(* IEC 61131-3 sources: volt/packages/volt-lsp-iec/test-corpus/awa-palletizer/Device/Plc Logic/Application/Library Manager/L_SEMP_ErrorManagement, 51 files *)

(* ---- EVTPARAM_CMPLENZEERRORMANAGEMENTACCESSACTSTATEDETERMINEEVENTCHANGED.dut ---- *)
TYPE EVTPARAM_CMPLENZEERRORMANAGEMENTACCESSACTSTATEDETERMINEEVENTCHANGED :
STRUCT
	SEVERITY : USINT;
	EVENTID : WORD;
	TEXTREFID : WORD;
	ACTSTATEDETERMINEEVENT : DWORD;
END_STRUCT
END_TYPE

(* ---- EVTPARAM_CMPLENZEERRORMANAGEMENTACCESSACTSTATEDETERMINEEVENTCHANGED_V2.dut ---- *)
TYPE EVTPARAM_CMPLENZEERRORMANAGEMENTACCESSACTSTATEDETERMINEEVENTCHANGED_V2 :
STRUCT
	SEVERITY : USINT;
	EVENTID : WORD;
	TEXTREFID : WORD;
	ACTSTATEDETERMINEEVENT : DWORD;
	USERGROUP : WORD;
	USERPRIORITY : WORD;
	EVENTCONTROL : WORD;
END_STRUCT
END_TYPE

(* ---- EVTPARAM_CMPLENZEERRORMANAGEMENTACCESSCOMMANDEVENTREACTION.dut ---- *)
TYPE EVTPARAM_CMPLENZEERRORMANAGEMENTACCESSCOMMANDEVENTREACTION :
STRUCT
	SEVERITY : USINT;
	EVENTID : WORD;
	TEXTREFID : WORD;
END_STRUCT
END_TYPE

(* ---- EVTPARAM_CMPLENZEERRORMANAGEMENTACCESSRESETCOMPONENTOCCURRED.dut ---- *)
TYPE EVTPARAM_CMPLENZEERRORMANAGEMENTACCESSRESETCOMPONENTOCCURRED :
STRUCT
	INSTANCEID : UDINT;
	LAYER : USINT;
	SEVERITY : USINT;
	STATE : USINT;
	EVENTID : WORD;
	TEXTREFID : WORD;
END_STRUCT
END_TYPE

(* ---- EVTPARAM_CMPLENZEERRORMANAGEMENTACCESSRESETOCCURRED.dut ---- *)
TYPE EVTPARAM_CMPLENZEERRORMANAGEMENTACCESSRESETOCCURRED :
STRUCT
	ACTHIGHESTPRIOREVENT : POINTER TO L_SEMP_ActEvent;
	PCOMPLIST : POINTER TO L_SEMP_ComponentListResetOccured;
END_STRUCT
END_TYPE

(* ---- L_SEMP_ACTEVENT.dut ---- *)
TYPE L_SEMP_ACTEVENT :
STRUCT
	LAYER : USINT;
	SEVERITY : USINT;
	STATE : USINT;
	EVENTID : WORD;
	TEXTREFID : WORD;
	INSTANCEID : DWORD;
	ACTSTATEDETERMINEEVENT : DWORD;
	TIMESTAMP : L_SEMP_LogTimeStamp;
END_STRUCT
END_TYPE

(* ---- L_SEMP_BEHAVIOUR.dut ---- *)
TYPE L_SEMP_BEHAVIOUR :
(
	PROCESSERRORREACTION := 0,
	ONLYLOGGING := 1
);
END_TYPE

(* ---- L_SEMP_COMPONENTLISTRESETOCCURED.dut ---- *)
TYPE L_SEMP_COMPONENTLISTRESETOCCURED :
STRUCT
	PREVCMP : POINTER TO L_SEMP_ComponentListResetOccured;
	PCOMPONENT : POINTER TO DWORD;
	NEXTCMP : POINTER TO L_SEMP_ComponentListResetOccured;
END_STRUCT
END_TYPE

(* ---- L_SEMP_EVENTCONTROL.dut ---- *)
TYPE L_SEMP_EVENTCONTROL :
(
	NOACKNOLAGENEEDED := 0,
	ACKNOLAGENEEDED := 1,
	EVENTCONTROLNOTUSED := 255
);
END_TYPE

(* ---- L_SEMP_EVENTPARAMETERS.dut ---- *)
TYPE L_SEMP_EVENTPARAMETERS :
STRUCT
	EVENTPARAMETERS : ARRAY [1..10] OF L_SEMP_ParameterItem;
END_STRUCT
END_TYPE

(* ---- L_SEMP_EVENTPARAMETERSSHORT.dut ---- *)
TYPE L_SEMP_EVENTPARAMETERSSHORT :
STRUCT
	EVENTPARAMETERS : ARRAY [1..10] OF L_SEMP_ParameterItemShort;
END_STRUCT
END_TYPE

(* ---- L_SEMP_GROUP.dut ---- *)
TYPE L_SEMP_GROUP :
(
	USERGROUP1 := 1,
	USERGROUP2 := 2,
	USERGROUP3 := 3,
	USERGROUP4 := 4,
	USERGROUP5 := 5,
	MANUFACTURERGROUP1 := 11,
	MANUFACTURERGROUP2 := 12
);
END_TYPE

(* ---- L_SEMP_LAYER.dut ---- *)
TYPE L_SEMP_LAYER :
(
	KINEMATICS := 6,
	MOTION := 7,
	APPLICATION := 8,
	IEC_APPLICATION := 40,
	TA_LAYER := 50
);
END_TYPE

(* ---- L_SEMP_LAYER_INTERN.dut ---- *)
TYPE L_SEMP_LAYER_INTERN :
(
	LEM_LA_I900_BASE_FW := 0,
	LEM_LA_SAFETY := 1,
	LEM_LA_FEEDBACK := 2,
	LEM_LA_ETC_SLAVE := 3,
	LEM_LA_BASE_SETTINGS := 4,
	LEM_LA_COMMUNICATION := 5,
	LEM_LA_KINEMATICS := 6,
	LEM_LA_MOTION := 7,
	LEM_LA_TECH_APPLICATION := 8,
	LEM_LA_FIELDBUS := 10,
	LEM_LA_LEM := 20,
	LEM_LA_IEC_RUNTIME := 30,
	LEM_LA_ETC_MASTER := 31,
	LEM_LA_I900_IO_DRIVER := 32,
	LEM_LA_IEC_APPLICATION := 40,
	LEM_LA_TA_LAYER := 50
);
END_TYPE

(* ---- L_SEMP_LOGTIMESTAMP.dut ---- *)
TYPE L_SEMP_LOGTIMESTAMP :
STRUCT
	DWLOWDATETIME : DWORD;
	DWHIGHDATETIME : DWORD;
END_STRUCT
END_TYPE

(* ---- L_SEMP_PARAMETERITEM.dut ---- *)
TYPE L_SEMP_PARAMETERITEM :
STRUCT
	SIZE : BYTE;
	ETYPE : INT;
	VALUE : L_SEMP_ParaValue;
END_STRUCT
END_TYPE

(* ---- L_SEMP_PARAMETERITEMSHORT.dut ---- *)
TYPE L_SEMP_PARAMETERITEMSHORT :
STRUCT
	SIZE : BYTE;
	ETYPE : INT;
	VALUE : L_SEMP_ParaValueShort;
END_STRUCT
END_TYPE

(* ---- L_SEMP_PARAVALUE.dut ---- *)
TYPE L_SEMP_PARAVALUE :
UNION
	DWVALUE : DWORD;
	DNVALUE : DINT;
	FVALUE : REAL;
	STVALUE : STRING;
	DWTEXTLISTID : DWORD;
END_UNION
END_TYPE

(* ---- L_SEMP_PARAVALUESHORT.dut ---- *)
TYPE L_SEMP_PARAVALUESHORT :
UNION
	DWVALUE : DWORD;
	DNVALUE : DINT;
	RVALUE : REAL;
	LRVALUE : LREAL;
	DWTEXTLISTID : DWORD;
END_UNION
END_TYPE

(* ---- L_SEMP_PRIORITY.dut ---- *)
TYPE L_SEMP_PRIORITY :
(
	PRIORITY_1 := 1,
	PRIORITY_2 := 2,
	PRIORITY_3 := 3,
	PRIORITY_4 := 4,
	PRIORITY_5 := 5,
	PRIORITY_INFO_NOT_USED := 255
);
END_TYPE

(* ---- L_SEMP_SERVERITY.dut ---- *)
TYPE L_SEMP_SERVERITY :
(
	LEM_SEV_NO_RESPONSE := 0,
	LEM_SEV_FAULT_CIA402 := 1,
	LEM_SEV_WARNING := 2,
	LEM_SEV_INFORMATION := 11,
	LEM_SEV_WARNING_LOCK := 13,
	LEM_SEV_TROUBLE_LOG := 15,
	LEM_SEV_TROUBLE := 16,
	LEM_SEV_FAULT_LOG := 18,
	LEM_SEV_FAULT_FAST_STOP := 19,
	LEM_SEV_FAULT_QSP := 20,
	LEM_SEV_FAULT_CINH := 21,
	LEM_SEV_FAULT := 23
);
END_TYPE

(* ---- L_SEMP_SERVERITYLEVEL.dut ---- *)
TYPE L_SEMP_SERVERITYLEVEL :
(
	NO_RESPONSE := 0,
	FAULT_CIA402 := 1,
	WARNING := 2,
	INFORMATION := 11,
	WARNING_LOCK := 13,
	TROUBLE_LOG := 15,
	TROUBLE := 16,
	FAULT_FAST_STOP := 19,
	FAULT_QSP := 20,
	FAULT_QSP_CINH := 21,
	FAULT := 23
);
END_TYPE

(* ---- L_SEMP_EVENTIDS.gvl ---- *)
VAR_GLOBAL
	CMPID_CMPLENZEERRORMANAGEMENTACCESS : DWORD := 16#2014;
	EVT_CMPLENZEERRORMANAGEMENTACCESSACTSTATEDETERMINEEVENTCHANGED : DWORD := 16#10000011;
	EVTPARAMID_CMPLENZEERRORMANAGEMENTACCESSACTSTATEDETERMINEEVENTCHANGED : WORD := 16#1;
	EVTVERSION_CMPLENZEERRORMANAGEMENTACCESSACTSTATEDETERMINEEVENTCHANGED : WORD := 16#1;
	EVT_CMPLENZEERRORMANAGEMENTACCESSRESETOCCURRED : DWORD := 16#10000012;
	EVTPARAMID_CMPLENZEERRORMANAGEMENTACCESSRESETOCCURRED : WORD := 16#1;
	EVTVERSION_CMPLENZEERRORMANAGEMENTACCESSRESETOCCURRED : WORD := 16#1;
	EVT_CMPLENZEERRORMANAGEMENTACCESSCOMMANDEVENTREACTION : DWORD := 16#10000013;
	EVTPARAMID_CMPLENZEERRORMANAGEMENTACCESSCOMMANDEVENTREACTION : WORD := 16#1;
	EVTVERSION_CMPLENZEERRORMANAGEMENTACCESSCOMMANDEVENTREACTION : WORD := 16#1;
	EVT_CMPLENZEERRORMANAGEMENTACCESSREADACTERRORDATAAVAILABLE : DWORD := 16#10000014;
	EVTPARAMID_CMPLENZEERRORMANAGEMENTACCESSREADACTERRORDATAAVAILABLE : WORD := 16#1;
	EVTVERSION_CMPLENZEERRORMANAGEMENTACCESSREADACTERRORDATAAVAILABLE : WORD := 16#1;
END_VAR

(* ---- GETBOOLEANPROPERTY.pou ---- *)
FUNCTION GETBOOLEANPROPERTY : BOOL
VAR_INPUT
	STKEY : WSTRING;
END_VAR
END_FUNCTION

(* ---- GETCOMPANY.pou ---- *)
FUNCTION GETCOMPANY : WSTRING
END_FUNCTION

(* ---- GETNUMBERPROPERTY.pou ---- *)
FUNCTION GETNUMBERPROPERTY : DINT
VAR_INPUT
	STKEY : WSTRING;
END_VAR
END_FUNCTION

(* ---- GETTEXTPROPERTY.pou ---- *)
FUNCTION GETTEXTPROPERTY : WSTRING
VAR_INPUT
	STKEY : WSTRING;
END_VAR
END_FUNCTION

(* ---- GETTEXTPROPERTY2.pou ---- *)
FUNCTION GETTEXTPROPERTY2 : POINTER TO WSTRING
VAR_INPUT
	STKEY : WSTRING;
END_VAR
END_FUNCTION

(* ---- GETTITLE.pou ---- *)
FUNCTION GETTITLE : WSTRING
END_FUNCTION

(* ---- GETVERSION.pou ---- *)
FUNCTION GETVERSION : VERSION
END_FUNCTION

(* ---- GETVERSIONPROPERTY.pou ---- *)
FUNCTION GETVERSIONPROPERTY : VERSION
VAR_INPUT
	STKEY : WSTRING;
END_VAR
END_FUNCTION

(* ---- L_SEMP_CLEAREVENT.pou ---- *)
FUNCTION L_SEMP_CLEAREVENT : RTS_IEC_RESULT
VAR_INPUT
	HHANDLE : RTS_IEC_HANDLE := RTS_INVALID_HANDLE;
	UIEVENTID : UINT := 16#0;
END_VAR
END_FUNCTION

(* ---- L_SEMP_CLEAREVENT_V2.pou ---- *)
FUNCTION L_SEMP_CLEAREVENT_V2 : RTS_IEC_RESULT
VAR_INPUT
	HHANDLE : RTS_IEC_HANDLE := RTS_INVALID_HANDLE;
	UIEVENTID : UINT := 16#0;
	UITEXTREFID : UINT := 16#0;
END_VAR
END_FUNCTION

(* ---- L_SEMP_GETACCESSACTSTATEDETERMINEPARAMETER.pou ---- *)
FUNCTION L_SEMP_GETACCESSACTSTATEDETERMINEPARAMETER : BOOL
VAR_INPUT
	PPARAMETER : POINTER TO BYTE;
	SEVERITY : POINTER TO USINT;
	EVENTID : POINTER TO WORD;
	TEXTREFID : POINTER TO WORD;
	ACTSTATEDETERMINEEVENT : POINTER TO DWORD;
END_VAR
END_FUNCTION

(* ---- L_SEMP_GETACCESSACTSTATEDETERMINEPARAMETER2.pou ---- *)
FUNCTION L_SEMP_GETACCESSACTSTATEDETERMINEPARAMETER2 : BOOL
VAR_INPUT
	PPARAMETER : POINTER TO BYTE;
	SEVERITY : POINTER TO USINT;
	EVENTID : POINTER TO WORD;
	TEXTREFID : POINTER TO WORD;
	ACTSTATEDETERMINEEVENT : POINTER TO DWORD;
	ACTERRORCODE : POINTER TO DWORD;
END_VAR
END_FUNCTION

(* ---- L_SEMP_GETACCESSACTSTATEDETERMINEPARAMETER3.pou ---- *)
FUNCTION L_SEMP_GETACCESSACTSTATEDETERMINEPARAMETER3 : BOOL
VAR_INPUT
	PPARAMETER : POINTER TO BYTE;
	SEVERITY : POINTER TO USINT;
	EVENTID : POINTER TO WORD;
	TEXTREFID : POINTER TO WORD;
	ACTSTATEDETERMINEEVENT : POINTER TO DWORD;
	ACTERRORCODE : POINTER TO DWORD;
	USERGROUP : POINTER TO USINT;
END_VAR
END_FUNCTION

(* ---- L_SEMP_GETCOMMANDEVENTREACTIONPARAMETER.pou ---- *)
FUNCTION L_SEMP_GETCOMMANDEVENTREACTIONPARAMETER : BOOL
VAR_INPUT
	PPARAMETER : POINTER TO BYTE;
	SEVERITY : POINTER TO USINT;
	EVENTID : POINTER TO WORD;
	TEXTREFID : POINTER TO WORD;
END_VAR
END_FUNCTION

(* ---- L_SEMP_GETRESETOCUREDINCOMPONENT.pou ---- *)
FUNCTION L_SEMP_GETRESETOCUREDINCOMPONENT : BOOL
VAR_INPUT
	PPARAMETER : POINTER TO BYTE;
	PCOMPONENT : POINTER TO DWORD;
	PACTSEVERITY : POINTER TO USINT;
END_VAR
END_FUNCTION

(* ---- L_SEMP_NOTIFYEVENT.pou ---- *)
FUNCTION L_SEMP_NOTIFYEVENT : RTS_IEC_RESULT
VAR_INPUT
	HHANDLE : RTS_IEC_HANDLE := RTS_INVALID_HANDLE;
	UIEVENTID : UINT := 16#0;
	ESEVERITY : L_SEMP_Serverity := L_SEMP_Serverity.LEM_SEV_NO_RESPONSE;
	UITEXTREFID : UINT := 16#0;
	UINUMPARAM : UINT := 16#0;
	PPARAMETES : POINTER TO L_SEMP_EventParameters;
END_VAR
END_FUNCTION

(* ---- L_SEMP_NOTIFYEVENT_V2.pou ---- *)
FUNCTION L_SEMP_NOTIFYEVENT_V2 : RTS_IEC_RESULT
VAR_INPUT
	HHANDLE : RTS_IEC_HANDLE := RTS_INVALID_HANDLE;
	UIEVENTID : UINT := 16#0;
	ESEVERITY : USINT := L_SEMP_Serverity.LEM_SEV_NO_RESPONSE;
	UITEXTREFID : UINT := 16#0;
	UINUMPARAM : UINT := 16#0;
	PPARAMETES : POINTER TO L_SEMP_EventParameters;
	UIEVENTCONTROL : UINT := 16#0;
	UIUSERPRIORITY : UINT := 16#0;
	UITARGETGROUP : UINT := 16#0;
END_VAR
END_FUNCTION

(* ---- L_SEMP_NOTIFYEVENTSHORT.pou ---- *)
FUNCTION L_SEMP_NOTIFYEVENTSHORT : RTS_IEC_RESULT
VAR_INPUT
	HHANDLE : RTS_IEC_HANDLE := RTS_INVALID_HANDLE;
	UIEVENTID : UINT := 16#0;
	ESEVERITY : L_SEMP_Serverity := L_SEMP_Serverity.LEM_SEV_NO_RESPONSE;
	UITEXTREFID : UINT := 16#0;
	UINUMPARAM : UINT := 16#0;
	PPARAMETES : POINTER TO L_SEMP_EventParametersShort;
END_VAR
END_FUNCTION

(* ---- L_SEMP_NOTIFYEVENTSHORT_V2.pou ---- *)
FUNCTION L_SEMP_NOTIFYEVENTSHORT_V2 : RTS_IEC_RESULT
VAR_INPUT
	HHANDLE : RTS_IEC_HANDLE := RTS_INVALID_HANDLE;
	UIEVENTID : UINT := 16#0;
	ESEVERITY : L_SEMP_Serverity := L_SEMP_Serverity.LEM_SEV_NO_RESPONSE;
	UITEXTREFID : UINT := 16#0;
	UINUMPARAM : UINT := 16#0;
	PPARAMETES : POINTER TO L_SEMP_EventParametersShort;
	UIEVENTCONTROL : UINT := 16#0;
	UIUSERPRIORITY : UINT;
	UITARGETGROUP : UINT := 16#0;
END_VAR
END_FUNCTION

(* ---- L_SEMP_NOTIFYEVENTSHORT_V3.pou ---- *)
FUNCTION L_SEMP_NOTIFYEVENTSHORT_V3 : RTS_IEC_RESULT
VAR_INPUT
	HHANDLE : RTS_IEC_HANDLE := RTS_INVALID_HANDLE;
	UIEVENTID : UINT := 16#0;
	ESEVERITY : L_SEMP_Serverity := L_SEMP_Serverity.LEM_SEV_NO_RESPONSE;
	UITEXTREFID : UINT := 16#0;
	UINUMPARAM : UINT := 16#0;
	PPARAMETES : POINTER TO L_SEMP_EventParametersShort;
	UIEVENTCONTROL : UINT := 16#0;
	UIREACTION : UINT := 0;
	UITARGETGROUP : UINT := 16#0;
END_VAR
END_FUNCTION

(* ---- L_SEMP_REGISTERCOMPONENT.pou ---- *)
FUNCTION L_SEMP_REGISTERCOMPONENT : RTS_IEC_HANDLE
VAR_INPUT
	SCOMPONENTNAME : STRING := '';
	UILAYER : UINT := 16#0;
	UITEXTREFID : UINT := 16#0;
	UIREAKTIONITF : UINT := 16#0;
END_VAR
END_FUNCTION

(* ---- L_SEMP_REGISTERCOMPONENT2.pou ---- *)
FUNCTION L_SEMP_REGISTERCOMPONENT2 : RTS_IEC_HANDLE
VAR_INPUT
	SCOMPONENTNAME : STRING := '';
	UILAYER : UINT := 16#0;
	UITEXTREFID : UINT := 16#0;
	UIREAKTIONITF : UINT := 16#0;
	UIGETALLRESETS : UINT := 16#0;
END_VAR
END_FUNCTION

(* ---- L_SEMP_REQUESTRESET.pou ---- *)
FUNCTION L_SEMP_REQUESTRESET : RTS_IEC_RESULT
VAR_INPUT
	HHANDLE : RTS_IEC_HANDLE := RTS_INVALID_HANDLE;
END_VAR
END_FUNCTION

(* ---- L_SEMP_REQUESTRESETCOMPONENT.pou ---- *)
FUNCTION L_SEMP_REQUESTRESETCOMPONENT : RTS_IEC_RESULT
VAR_INPUT
	HHANDLE : RTS_IEC_HANDLE := RTS_INVALID_HANDLE;
END_VAR
END_FUNCTION

(* ---- L_SEMP_REQUESTRESETCOMPONENTLIST.pou ---- *)
FUNCTION L_SEMP_REQUESTRESETCOMPONENTLIST : RTS_IEC_RESULT
VAR_INPUT
	HANDLELIST : POINTER TO RTS_IEC_HANDLE;
	LISTCOUNT : WORD;
END_VAR
END_FUNCTION

(* ---- L_SEMP_UNREGISTERCOMPONENT.pou ---- *)
FUNCTION L_SEMP_UNREGISTERCOMPONENT : RTS_IEC_RESULT
VAR_INPUT
	HHANDLE : RTS_IEC_HANDLE := RTS_INVALID_HANDLE;
END_VAR
END_FUNCTION

(* ---- L_SEMP_READACTUALERRORCODE.pou ---- *)
FUNCTION_BLOCK L_SEMP_READACTUALERRORCODE
VAR_INPUT
	XENABLE : BOOL;
END_VAR
VAR_OUTPUT
	XBUSY : BOOL;
	DWERRORCODE : DWORD;
	ESEVERITY : L_SEMP_ServerityLevel;
END_VAR
VAR
	ITFCALLBACK : CmpEventMgr.ICmpEventCallback;
	HEVENTUPDATEACTIVEERROR : RTS_IEC_HANDLE := SysTypes.RTS_INVALID_HANDLE;
	HINTERFACEUPDATEACTIVEERROR : RTS_IEC_HANDLE := SysTypes.RTS_INVALID_HANDLE;
	WEVTCOUNT_UPDATEACTIVEERROR : WORD;
	SEVERITY_INT : USINT;
	EVENTID_INT : WORD;
	USERGROUP_INT : USINT;
	EUSERGROUP : USINT;
	TEXTREFID_INT : WORD;
	ACTSTATEDETERMINEEVENT_INT : DWORD;
	ACTERRORCODE_INT : DWORD;
	USERGROUP : USINT;
END_VAR
END_FUNCTION_BLOCK

METHOD FB_EXIT : BOOL
VAR_INPUT
	BINCOPYCODE : BOOL;
END_VAR
END_METHOD

METHOD FB_INIT : BOOL
VAR_INPUT
	BINITRETAINS : BOOL;
	BINCOPYCODE : BOOL;
END_VAR
END_METHOD

METHOD EVENTCALLBACK : UDINT
VAR_INPUT
	PEVENTPARAM : POINTER TO EventParam;
END_VAR
END_METHOD

METHOD REGISTEREVENT
END_METHOD

METHOD UNREGISTEREVENT
END_METHOD

(* ---- L_SEMP_SETERROR.pou ---- *)
FUNCTION_BLOCK L_SEMP_SETERROR
VAR_INPUT
	XRESETERROR : BOOL;
	XSETERROR1 : BOOL;
	ESEVERITY1 : L_SEMP_ServerityLevel;
	WERRORID1 : WORD;
	WTEXTREFID1 : WORD;
	XSETERROR2 : BOOL;
	ESEVERITY2 : L_SEMP_ServerityLevel;
	WERRORID2 : WORD;
	WTEXTREFID2 : WORD;
	XSETERROR3 : BOOL;
	ESEVERITY3 : L_SEMP_ServerityLevel;
	WERRORID3 : WORD;
	WTEXTREFID3 : WORD;
	XSETERROR4 : BOOL;
	ESEVERITY4 : L_SEMP_ServerityLevel;
	WERRORID4 : WORD;
	WTEXTREFID4 : WORD;
END_VAR
VAR_OUTPUT
	XERROR : BOOL;
	EERRORID : L_IE1P_Error;
	XERRORRESETACTIVE : BOOL;
END_VAR
VAR
	ERRORHANDLE : RTS_IEC_HANDLE := 0;
	ELAYER : L_SEMP_Layer := L_SEMP_Layer.Application;
	EERRORBEHAVIOUR : L_SEMP_Behaviour := L_SEMP_Behaviour.ProcessErrorReaction;
	SCOMPONENTNAME : STRING := '';
	WDEFAULTTEXTREFID : WORD := 16#2C00;
	XDEFAULTTEXTREFIDVALID : BOOL;
	XRESETERROROLD : BOOL;
	XSETERROR1OLD : BOOL;
	XSETERROR2OLD : BOOL;
	XSETERROR3OLD : BOOL;
	XSETERROR4OLD : BOOL;
	SINSTANCESTR : STRING;
	SINSTANCESTRDUMMY : STRING;
	ESEVERITY1_INT : L_SEMP_ServerityLevel;
	ESEVERITY2_INT : L_SEMP_ServerityLevel;
	ESEVERITY3_INT : L_SEMP_ServerityLevel;
	ESEVERITY4_INT : L_SEMP_ServerityLevel;
	WERRORID1_INT : WORD;
	WERRORID2_INT : WORD;
	WERRORID3_INT : WORD;
	WERRORID4_INT : WORD;
	ITFCALLBACK : CmpEventMgr.ICmpEventCallback;
	HEVENTRESETOCCURED : RTS_IEC_HANDLE := SysTypes.RTS_INVALID_HANDLE;
	HINTERFACERESETOCCURED : RTS_IEC_HANDLE := SysTypes.RTS_INVALID_HANDLE;
	WEVTCOUNT_RESETOCCURED : WORD;
	XRESETOCCURED : BOOL;
	XFBERRORINT1 : BOOL;
	EFBERRORIDINT1 : L_IE1P_Error;
	XFBERRORINT2 : BOOL;
	EFBERRORIDINT2 : L_IE1P_Error;
	XFBERRORINT3 : BOOL;
	EFBERRORIDINT3 : L_IE1P_Error;
	XFBERRORINT4 : BOOL;
	EFBERRORIDINT4 : L_IE1P_Error;
	COMPONENTNAME : STRING;
	DEFAULTTEXTREFID : WORD;
	ERRORBEHAVIOUR : L_SEMP_Behaviour;
	LAYER : L_SEMP_Layer;
END_VAR
END_FUNCTION_BLOCK

METHOD CHECKSETERROR : STRING
VAR_IN_OUT
	XSETERROR : BOOL;
	XSETERROROLD : BOOL;
	ESEVERITY : L_SEMP_Serverity;
	ESEVERITY_INT : L_SEMP_Serverity;
	WERRORID : WORD;
	WERRORID_INT : WORD;
	WTEXTREFID : WORD;
	XFBERRORINT : BOOL;
	EFBERRORIDINT : L_IE1P_Error;
END_VAR
END_METHOD

METHOD GETINSTANCENAME : STRING
END_METHOD

METHOD FB_AFTERINIT
END_METHOD

METHOD FB_EXIT : BOOL
VAR_INPUT
	BINCOPYCODE : BOOL;
END_VAR
END_METHOD

METHOD FB_INIT : BOOL
VAR_INPUT
	BINITRETAINS : BOOL;
	BINCOPYCODE : BOOL;
END_VAR
END_METHOD

METHOD EVENTCALLBACK : UDINT
VAR_INPUT
	PEVENTPARAM : POINTER TO EventParam;
END_VAR
END_METHOD

METHOD REGISTEREVENT
END_METHOD

METHOD UNREGISTEREVENT
END_METHOD
